{attribute 'qualified_only'}
{attribute 'strict'}
{attribute 'to_string'}
TYPE E_LWord :
(
	eOptionA := 0,
	eOptionB,
	eOptionC
) LWORD;
END_TYPE

(* stored: Version 1.1.0.1, ProductVersion 3.1.4026.19
   DUT E_LWord: Id {f9196696-6b9f-4ab1-ad1c-f9bacb46f274} *)
